// TIA Portal V21 export
// export: Created 2026-11-11T00:48:12.3484958Z, ExportSetting WithDefaults, DisplayName Totally Integrated Automation Portal, DisplayVersion V21 Update 3, DisplayName STEP 7 Professional, DisplayVersion V21 Update 3, DisplayName STEP 7 Safety, DisplayVersion V21, DisplayName Tech WebApplication, DisplayVersion V21, DisplayName WinCC Basic/Comfort/Advanced, DisplayVersion V21 Update 3, DisplayName WinCC Unified, DisplayVersion V21 Update 3
FUNCTION_BLOCK "FB_Scl_sl026"   // FB40, SCL
{ S7_Optimized_Access := 'TRUE' }
VERSION : 0.1
// stored: AutoNumber true, IsIECCheckEnabled false, IsRetainMemResEnabled false, MemoryReserve 100, SetENOAutomatically false, UDAEnableTagReadback false
   VAR_INPUT
      v_in1 : Time;
      v_in2 : Time;
   END_VAR
   VAR_OUTPUT
      v_ret : Time;
   END_VAR
BEGIN
   #v_ret := MAX(IN1 := #v_in1, IN2 := #v_in2);
END_FUNCTION_BLOCK
